// TIA Portal V20 export
// export: Created 2026-10-12T16:46:21.3909461Z, ExportSetting WithDefaults, DisplayName Totally Integrated Automation Portal, DisplayVersion V20 Update 6, DisplayName TIA Portal Openness, DisplayVersion V20 Update 6, DisplayName TIA Portal Version Control Interface, DisplayVersion V20 Update 6, DisplayName SINAMICS Startdrive Advanced, DisplayVersion V20 SP1 Update 2, DisplayName SINAMICS Startdrive G110M, G120, G120C, G120D, G120P, G115D, DisplayVersion V20 SP1 Update 2, DisplayName SINAMICS Startdrive G130, G150, S120, S150, SINAMICS MV, G220, S200, S210, DisplayVersion V20 SP1 Update 2, DisplayName STEP 7 Professional, DisplayVersion V20 Update 6, DisplayName STEP 7 Safety, DisplayVersion V20 Update 2, DisplayName WinCC Basic/Comfort/Advanced, DisplayVersion V20 Update 6, DisplayName WinCC Professional, DisplayVersion V20 Update 6, DisplayName WinCC Unified, DisplayVersion V20 Update 6
DATA_BLOCK "FB_Auftragsmanager_DB"   // DB11
VERSION : 0.1
// stored: AutoNumber true, DBAccessibleFromOPCUA true, DBAccessibleFromWebserver true, InstanceOfName FB_Auftragsmanager, InstanceOfType FB
"FB_Auftragsmanager"
   // VAR_IN_OUT
   //    Auftraege : Array[0..9] of "UDT_Prozessroute";
   //    Bad_Konfig : Array[1.."c_Anzahl_Bad"] of "UDT_Bad_Konfig";
   // END_VAR
   // VAR
   //    Freigabe_Alt : Array[0..9] of Bool;
   // END_VAR
BEGIN
END_DATA_BLOCK
